% RSLogix 500 project PROGRAM 2.RSS, saved by version 8.30.00.16 %
PROJECT "UNTITLED"    % processor: Bul.1763 MicroLogix 1100 Series B %

PROGRAM FILES
  LAD 2 "MAIN"  3 rungs
  LAD 3 "IO"  8 rungs
  LAD 4 "PROC LOGIC"  11 rungs

DATA FILES
  O0 OUTPUT  4 elements
  I1 INPUT  6 elements
  S2 STATUS  66 elements
  B3 BINARY  2 elements
  T4 TIMER  1 elements
  C5 COUNTER  1 elements
  R6 CONTROL  1 elements
  N7 INTEGER  1 elements
  F8 FLOAT  1 elements

LADDER 2 "MAIN"
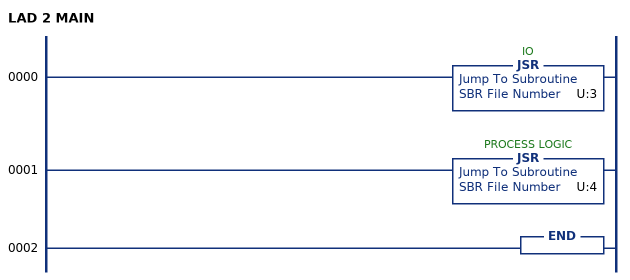
% Rung: 0 %
SOR JSR U:3 EOR
%   U:3  "IO" %
% Rung: 1 %
SOR JSR U:4 EOR
%   U:4  "PROCESS LOGIC" %
% Rung: 2 %
SOR END EOR

LADDER 3 "IO"
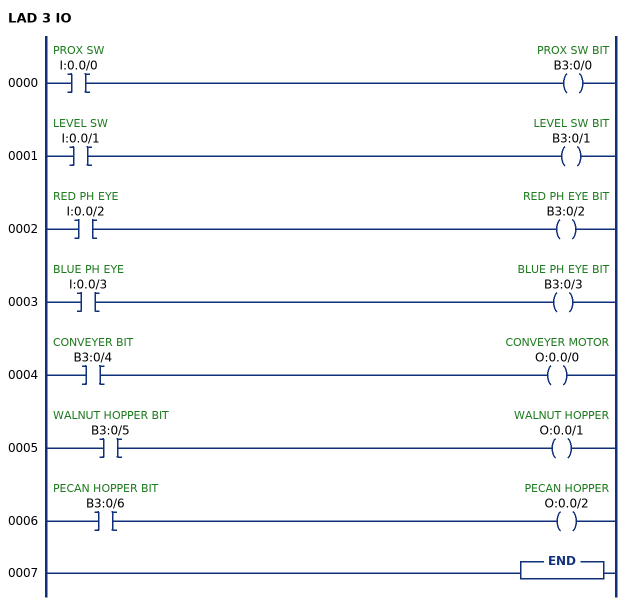
% Rung: 0 %
SOR XIC I:0.0/0 OTE B3:0/0 EOR
%   I:0.0/0  "PROX SW" %
%   B3:0/0  "PROX SW BIT" %
% Rung: 1 %
SOR XIC I:0.0/1 OTE B3:0/1 EOR
%   I:0.0/1  "LEVEL SW" %
%   B3:0/1  "LEVEL SW BIT" %
% Rung: 2 %
SOR XIC I:0.0/2 OTE B3:0/2 EOR
%   I:0.0/2  "RED PH EYE" %
%   B3:0/2  "RED PH EYE BIT" %
% Rung: 3 %
SOR XIC I:0.0/3 OTE B3:0/3 EOR
%   I:0.0/3  "BLUE PH EYE" %
%   B3:0/3  "BLUE PH EYE BIT" %
% Rung: 4 %
SOR XIC B3:0/4 OTE O:0.0/0 EOR
%   B3:0/4  "CONVEYER BIT" %
%   O:0.0/0  "CONVEYER MOTOR" %
% Rung: 5 %
SOR XIC B3:0/5 OTE O:0.0/1 EOR
%   B3:0/5  "WALNUT HOPPER BIT" %
%   O:0.0/1  "WALNUT HOPPER" %
% Rung: 6 %
SOR XIC B3:0/6 OTE O:0.0/2 EOR
%   B3:0/6  "PECAN HOPPER BIT" %
%   O:0.0/2  "PECAN HOPPER" %
% Rung: 7 %
SOR END EOR

LADDER 4 "PROC LOGIC"
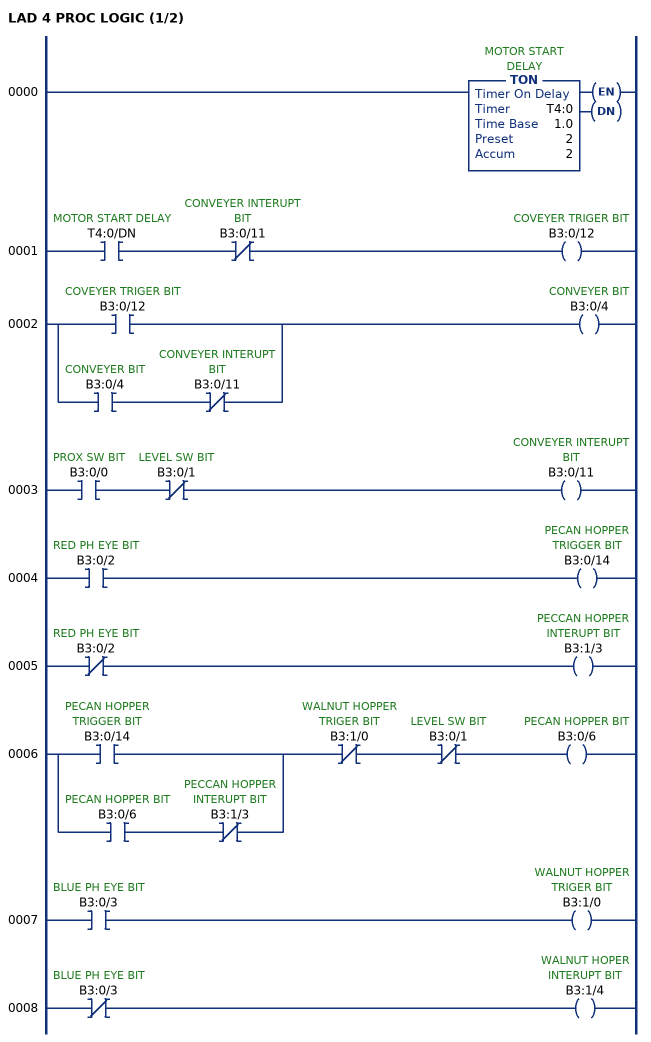
% Rung: 0 %
SOR TON T4:0 1.0 2 2 EOR
%   T4:0  "MOTOR START DELAY" %
% Rung: 1 %
SOR XIC T4:0/DN XIO B3:0/11 OTE B3:0/12 EOR
%   T4:0  "MOTOR START DELAY" %
%   B3:0/11  "CONVEYER INTERUPT BIT" %
%   B3:0/12  "COVEYER TRIGER BIT" %
% Rung: 2 %
SOR BST XIC B3:0/12 NXB XIC B3:0/4 XIO B3:0/11 BND OTE B3:0/4 EOR
%   B3:0/12  "COVEYER TRIGER BIT" %
%   B3:0/4  "CONVEYER BIT" %
%   B3:0/11  "CONVEYER INTERUPT BIT" %
% Rung: 3 %
SOR XIC B3:0/0 XIO B3:0/1 OTE B3:0/11 EOR
%   B3:0/0  "PROX SW BIT" %
%   B3:0/1  "LEVEL SW BIT" %
%   B3:0/11  "CONVEYER INTERUPT BIT" %
% Rung: 4 %
SOR XIC B3:0/2 OTE B3:0/14 EOR
%   B3:0/2  "RED PH EYE BIT" %
%   B3:0/14  "PECAN HOPPER TRIGGER BIT" %
% Rung: 5 %
SOR XIO B3:0/2 OTE B3:1/3 EOR
%   B3:0/2  "RED PH EYE BIT" %
%   B3:1/3  "PECCAN HOPPER INTERUPT BIT" %
% Rung: 6 %
SOR BST XIC B3:0/14 NXB XIC B3:0/6 XIO B3:1/3 BND XIO B3:1/0 XIO B3:0/1 OTE B3:0/6 EOR
%   B3:0/14  "PECAN HOPPER TRIGGER BIT" %
%   B3:0/6  "PECAN HOPPER BIT" %
%   B3:1/3  "PECCAN HOPPER INTERUPT BIT" %
%   B3:1/0  "WALNUT HOPPER TRIGER BIT" %
%   B3:0/1  "LEVEL SW BIT" %
% Rung: 7 %
SOR XIC B3:0/3 OTE B3:1/0 EOR
%   B3:0/3  "BLUE PH EYE BIT" %
%   B3:1/0  "WALNUT HOPPER TRIGER BIT" %
% Rung: 8 %
SOR XIO B3:0/3 OTE B3:1/4 EOR
%   B3:0/3  "BLUE PH EYE BIT" %
%   B3:1/4  "WALNUT HOPER INTERUPT BIT" %

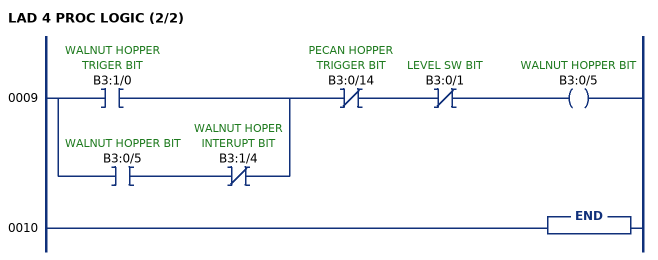
% Rung: 9 %
SOR BST XIC B3:1/0 NXB XIC B3:0/5 XIO B3:1/4 BND XIO B3:0/14 XIO B3:0/1 OTE B3:0/5 EOR
%   B3:1/0  "WALNUT HOPPER TRIGER BIT" %
%   B3:0/5  "WALNUT HOPPER BIT" %
%   B3:1/4  "WALNUT HOPER INTERUPT BIT" %
%   B3:0/14  "PECAN HOPPER TRIGGER BIT" %
%   B3:0/1  "LEVEL SW BIT" %
% Rung: 10 %
SOR END EOR

OTHER DOCUMENTED ADDRESSES
  B3:0/8  "CONVEYR MOTOR START BIT"
  B3:0/9  "ONS"
  B3:0/10  "ONS"
  B3:0/13  "ONS"
  B3:0/15  "ONS"
  B3:1/2  "ONS"
  T4:1  "MOTOR STOP DELAY"

DATA TABLE (non-zero values as saved)
DATA B3
% B3:0 % 0X466F 0X0005
DATA T4
% .PRE .ACC %
% T4:0 % 2 2
